// TIA Portal V21 export
// export: Created 2026-10-23T20:42:19.1657577Z, ExportSetting WithDefaults, DisplayName Totally Integrated Automation Portal, DisplayVersion V21 Update 1, DisplayName SINAMICS Startdrive Advanced, DisplayVersion V21 HF2, DisplayName SINAMICS Startdrive G110M, G120, G120C, G120D, G120P, G115D, DisplayVersion V21 HF2, DisplayName SINAMICS Startdrive G130, G150, S120, S150, G200, G220, S200, S210, S220, Innomotics MVD, DisplayVersion V21 HF2, DisplayName STEP 7 Professional, DisplayVersion V21 Update 1, DisplayName STEP 7 Safety, DisplayVersion V21, DisplayName Tech WebApplication, DisplayVersion V21, DisplayName WinCC Basic/Comfort/Advanced, DisplayVersion V21 Update 1, DisplayName WinCC Unified, DisplayVersion V21 Update 1
ORGANIZATION_BLOCK "OB_Cyclic100ms"   // OB35, SCL, CyclicInterrupt
TITLE = Weckalarm 100 ms / Cyclic interrupt 100 ms
{ S7_Optimized_Access := 'TRUE' }
VERSION : 0.1
// Ruft FB_SclTimers alle 100 ms mit eigener Instanz auf / Calls FB_SclTimers every 100 ms with its own instance
// stored: AutoNumber false, CyclicTime 100000, IsIECCheckEnabled false, PhaseOffset 20000, SetENOAutomatically false
   VAR_INPUT
      Initial_Call : Bool;   // Initial call of this OB
      Event_Count : Int;   // Events discarded
   END_VAR
BEGIN

       REGION Timers every 100 ms
           "IDB_SclTimersCyclic"(Start := "LevelHigh", Reset := "StopButton", DelayTime := T#1s);
       END_REGION

       REGION Analyzer C26l
           // The same instance is also called from OB_Main
           "IDB_AnaShared"(Pulse := "LevelHigh");
       END_REGION
END_ORGANIZATION_BLOCK
